Fanuc KAREL source: kx00002.compact.KL

PROGRAM KX00002
%STACKSIZE=65535
%PRIORITY=65535
%NOLOCKGROUP
VAR
I : INTEGER
J : INTEGER
B : BOOLEAN
F : FILE
S : STRING[80]
P : XYZWPR
BEGIN
OPEN FILE F ('RW','MD:KFSAMPLE.DT')
CLOSE FILE F
END KX00002
